PROGRAM RunSlave
VAR
	LampSlave_0: LampSlave;
	SlaveHandeshake_0: SlaveHandeshake;
	ixStrobOne :BOOL;
	ixStrobTwo :BOOL;
	startCar: BOOL;
	carEnd: BOOL;
	CarContorl_0: CarContorl;
END_VAR

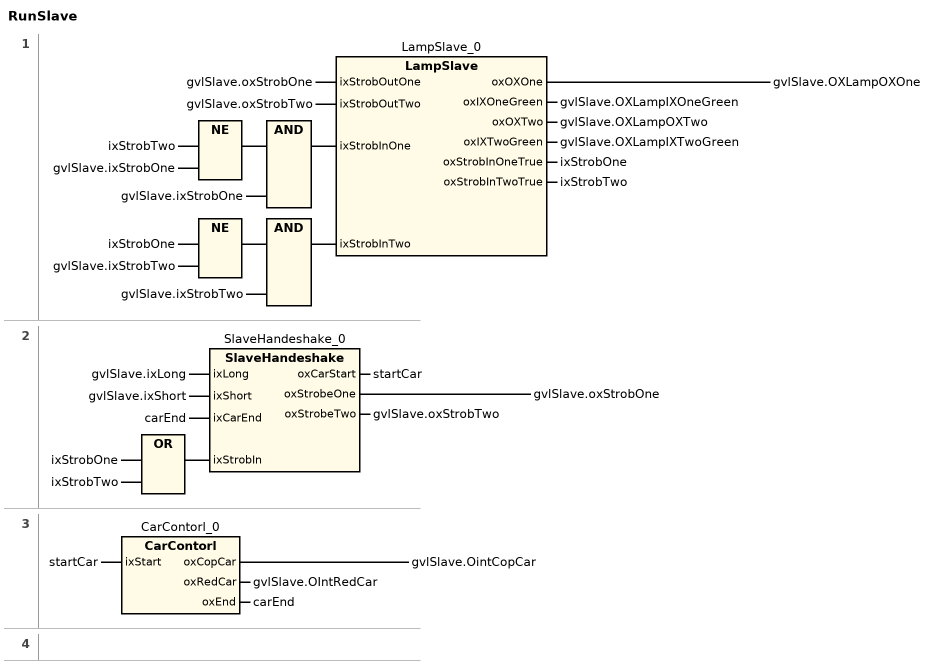
// NETWORK 1
LampSlave_0(
    ixStrobOutOne := gvlSlave.oxStrobOne,
    ixStrobOutTwo := gvlSlave.oxStrobTwo,
    ixStrobInOne := ixStrobTwo <> gvlSlave.ixStrobOne AND gvlSlave.ixStrobOne,
    ixStrobInTwo := ixStrobOne <> gvlSlave.ixStrobTwo AND gvlSlave.ixStrobTwo,
    oxIXOneGreen => gvlSlave.OXLampIXOneGreen,
    oxOXTwo => gvlSlave.OXLampOXTwo,
    oxIXTwoGreen => gvlSlave.OXLampIXTwoGreen,
    oxStrobInOneTrue => ixStrobOne,
    oxStrobInTwoTrue => ixStrobTwo); // LampSlave
gvlSlave.OXLampOXOne := LampSlave_0.oxOXOne;

// NETWORK 2
SlaveHandeshake_0(
    ixLong := gvlSlave.ixLong,
    ixShort := gvlSlave.ixShort,
    ixCarEnd := carEnd,
    ixStrobIn := ixStrobOne OR ixStrobTwo,
    oxCarStart => startCar,
    oxStrobeTwo => gvlSlave.oxStrobTwo); // SlaveHandeshake
gvlSlave.oxStrobOne := SlaveHandeshake_0.oxStrobeOne;

// NETWORK 3
CarContorl_0(ixStart := startCar, oxRedCar => gvlSlave.OIntRedCar, oxEnd => carEnd); // CarContorl
gvlSlave.OintCopCar := CarContorl_0.oxCopCar;

// NETWORK 4

END_PROGRAM

(* stored: Version 1.1.0.1, ProductVersion 3.1.4024.12
   POU RunSlave: Id {9d4154a5-7551-4a9b-be99-2aaf6aa886cb}, SpecialFunc None *)
